  OBJs.append(create_object_2(id=1, name="rack centrifuge", type=1, dimension=struct(length=0, width=0, height=0.106, diameter=0.020), gripper_offset=p[0,0,0.095,0,0,2.356]))
  OBJs.append(create_object_2(id=2, name="sample tube 1", type=2, dimension=struct(length=0, width=0, height=0.106, diameter=0.015), gripper_offset=p[0,0,0,0,0,0]))
  OBJs.append(create_object_2(id=3, name="rack sarstedt", type=3, dimension=struct(length=0, width=0, height=0.100, diameter=0.020), gripper_offset=p[0,0,0,0,0,0]))
  OBJs.append(create_object_2(id=4, name="Lab bottle", type=4, dimension=struct(length=0, width=0, height=0.100, diameter=0.030), gripper_offset=p[0,0,0.2,0,0,0]))
  def create_jig_2(id=0, name="", type=0, capacity=0, jig_offset=p[0,0,0,0,0,0]):
      # iformation about used jigs
      return struct(id=id, name=name, type=type, capacity=capacity, jig_offset=jig_offset)
  end

  JIG2 = create_jig_2()
  JIGs = make_list(0, create_jig_2(), 15)

  JIGs.append(create_jig_2(id=1, name="3FG", type=1, capacity=1, jig_offset=p[0,0,0,0,0,0]))
  JIGs.append(create_jig_2(id=2, name="jig input", type=2, capacity=1, jig_offset=p[0,0,0,0,0,-3.927]))
  JIGs.append(create_jig_2(id=3, name="jig output", type=3, capacity=1, jig_offset=p[0,0,0,0,0,0.78]))
  JIGs.append(create_jig_2(id=6, name="jig bin", type=6, capacity=1, jig_offset=p[0,0,0,0,0,0]))
  JIGs.append(create_jig_2(id=7, name="jig sarstedt racks", type=7, capacity=1, jig_offset=p[0,0,-0.02,0,0,0]))
  JIGs.append(create_jig_2(id=8, name="NoK Bin", type=8, capacity=1, jig_offset=p[0,0,0,0,0,0]))
  JIGs.append(create_jig_2(id=9, name="Pick bott jig", type=9, capacity=1, jig_offset=p[0,0,0,0,0,0]))
  JIGs.append(create_jig_2(id=10, name="Place bott jig", type=10, capacity=1, jig_offset=p[0,0,0,0,0,0]))
  JIGs.append(create_jig_2(id=11, name="bottle shake jig", type=11, capacity=1, jig_offset=p[0,0,0,0,0,0]))
  $ 20 "BeforeStarts"
  $ 21 "uLM"
  $ 22 "CMD_Stop≔ False "
  global CMD_Stop=  False
  $ 23 "CMD_Abort≔ False "
  global CMD_Abort=  False
  $ 24 "CMD_Clear≔ False "
  global CMD_Clear=  False
  $ 25 "STATE≔1"
  global STATE=1
  $ 26 "STATE_Info≔''"
  global STATE_Info=""
  $ 27 "ARM_Referenced≔ False "
  global ARM_Referenced=  False
  $ 28 "zero_ftsensor()"
  zero_ftsensor()
  $ 29 "poses init"
  $ 30 "PSE_A≔p[0,0,0,0,0,0]"
  global PSE_A=p[0,0,0,0,0,0]
  $ 31 "PSE_A_H≔p[0,0,0,0,0,0]"
  global PSE_A_H=p[0,0,0,0,0,0]
  $ 32 "PSE_R≔p[0,0,0,0,0,0]"
  global PSE_R=p[0,0,0,0,0,0]
  $ 33 "PSE_R_H≔p[0,0,0,0,0,0]"
  global PSE_R_H=p[0,0,0,0,0,0]
  $ 34 "PSE_T≔p[0,0,0,0,0,0]"
  global PSE_T=p[0,0,0,0,0,0]
  $ 35 "PSE_T_H≔p[0,0,0,0,0,0]"
  global PSE_T_H=p[0,0,0,0,0,0]
  $ 36 "PSE_C_E≔p[0,0,0,0,0,0]"
  global PSE_C_E=p[0,0,0,0,0,0]
  $ 37 "PSE_C_H≔p[0,0,0,0,0,0]"
  global PSE_C_H=p[0,0,0,0,0,0]
  $ 38 "PSE_C_S≔p[0,0,0,0,0,0]"
  global PSE_C_S=p[0,0,0,0,0,0]
  $ 39 "init_home_by_cartesian_pose(p[0,-0.400,0.300,0,0,0])"
  init_home_by_cartesian_pose(p[0,-0.400,0.300,0,0,0])
  $ 40 "Clearing"
  $ 41 "reset_error()"
  reset_error()
  $ 42 "reset_warning()"
  reset_warning()
  $ 43 "uGo"
  $ 45 "ugo_init( True ,'http://192.168.12.120:10001')"
  ugo_init(  True  ,"http://192.168.12.120:10001")
  $ 46 "ugo_update_outputs()"
  ugo_update_outputs()
  $ 47 "App"
  $ 48 "'ADD APPLICATION SPECIFIC COMMANDS'"
  # 'ADD APPLICATION SPECIFIC COMMANDS'
  $ 49 "Tools"
  $ 50 "OBJ_Picked≔gripper_has_object()"
  global OBJ_Picked=gripper_has_object()
  $ 51 "If OBJ_Picked"
  if (OBJ_Picked):
    # begin: URCap Program Node
    #   Source: Robotiq_Grippers, 1.8.4.4844, Robotiq Inc.
    #   Type: Gripper Activate
    $ 52 "Gripper Activate"

    kill rq_gripper_communication_thread
    rq_gripper_communication_thread_started = False

    rq_init_comm_if_connected(9, "1")
    rq_init_comm_if_connected(2, "2")
    rq_init_comm_if_connected(3, "3")
    rq_init_comm_if_connected(4, "4")
    rq_print_connected_grippers()
    rq_gripper_communication_thread = run rq_gripper_communication()

    while(not rq_gripper_communication_thread_started):
        sync()
    end

    rq_set_max_current_for_all_grippers()

    reset_and_activate = False

    rq_activate_all_grippers(False)
    # end: URCap Program Node
  else:
    $ 53 "Else" "noBreak"
    # begin: URCap Program Node
    #   Source: Robotiq_Grippers, 1.8.4.4844, Robotiq Inc.
    #   Type: Gripper Activate
    $ 54 "Gripper Reset and Activate"

    kill rq_gripper_communication_thread
    rq_gripper_communication_thread_started = False

    rq_init_comm_if_connected(9, "1")
    rq_init_comm_if_connected(2, "2")
    rq_init_comm_if_connected(3, "3")
    rq_init_comm_if_connected(4, "4")
    rq_print_connected_grippers()
    rq_gripper_communication_thread = run rq_gripper_communication()

    while(not rq_gripper_communication_thread_started):
        sync()
    end

    rq_set_max_current_for_all_grippers()

    reset_and_activate = True

    rq_activate_all_grippers(True)
    # end: URCap Program Node
  end
  $ 55 "zero_ftsensor()"
  zero_ftsensor()
  $ 56 "EXTT"
  $ 57 "Set GRP_3F_Enable=Off"
  set_standard_digital_out(4, False)
  $ 58 "Set GRP_3F_Decap=Off"
  set_standard_digital_out(3, False)
  $ 59 "Set GRP_3F_Cap=Off"
  set_standard_digital_out(2, False)
  $ 60 "Set GRP_3F_Open=Off"
  set_standard_digital_out(5, False)
  $ 61 "PSE_T≔get_tool_free_pose(dir=[0,0,0.150], move_in_base_frame=True)"
  global PSE_T=get_tool_free_pose(dir=[0,0,0.150], move_in_base_frame=True)
  $ 62 "If is_reachable(Base_const, [PSE_T])"
  if (is_reachable(p[0.0,0.0,0.0,0.0,0.0,0.0], [PSE_T])):
    $ 63 "MoveL"
    $ 64 "PSE_T" "breakAfter"
    movel(PSE_T, a=1.2, v=0.15)
  end
  while (True):
    $ 65 "Robot Program"
    $ 66 "MAIN"
    $ 67 "command_manager(external_control='uGO', cond_suspend=(ITM_Manipulated and AMR_AtTarget and AMR_Charging and AMR_Battery<40), cond_unsuspend=(AMR_Battery≟60))"
    command_manager(external_control="uGO", cond_suspend=(ITM_Manipulated  and  AMR_AtTarget  and  AMR_Charging  and  AMR_Battery<40), cond_unsuspend=(AMR_Battery == 60))
    $ 68 "log_state(STATE_Info)"
    log_state(STATE_Info)
    $ 69 "Switch STATE"
    switch_1 = STATE
    $ 70 "Case 1"
    if (1 == switch_1):
      $ 71 "Stopping"
      $ 72 "STATE_Info≔'Stopping'"
      global STATE_Info="Stopping"
      $ 73 "end_freedrive_mode()"
      end_freedrive_mode()
      $ 74 "Set"
      set_tcp(p[0.0,0.0,0.161,3.1415,0.0,0.0])
      $ 75 "PSE_T≔get_tool_free_pose(dir=[0,0,0.150], move_in_base_frame=True)"
      global PSE_T=get_tool_free_pose(dir=[0,0,0.150], move_in_base_frame=True)
      $ 76 "If is_reachable(Base_const, [PSE_T])"
      if (is_reachable(p[0.0,0.0,0.0,0.0,0.0,0.0], [PSE_T])):
        $ 77 "MoveL"
        $ 78 "PSE_T" "breakAfter"
        movel(PSE_T, a=1.2, v=0.15)
      end
      $ 79 "do_transition(keep_rxry=OBJ_Picked, r=0)"
      do_transition(keep_rxry=OBJ_Picked, r=0)
      $ 88 "Call Sub_AMR_MiR_V3"
      Sub_AMR_MiR_V3()
      $ 89 "If stopping() and AMR_Done"
      if (stopping()  and  AMR_Done):
        $ 90 "STATE≔2"
        global STATE=2
        $ 91 "ugo_update_outputs()"
        ugo_update_outputs()
      end
    elif (2 == switch_1):
      $ 92 "Case 2"
      $ 93 "Stopped"
      $ 94 "STATE_Info≔'Stopped'"
      global STATE_Info="Stopped"
      $ 95 "Call Sub_AMR_MiR_V3"
      Sub_AMR_MiR_V3()
      $ 96 "If CMD_Reset"
      if (CMD_Reset):
        $ 97 "STATE≔3"
        global STATE=3
        $ 98 "ugo_update_outputs()"
        ugo_update_outputs()
      end
    elif (3 == switch_1):
      $ 99 "Case 3"
      $ 100 " Resetting"
      $ 101 "STATE_Info≔'Resetting'"
      global STATE_Info="Resetting"
      $ 102 "uML"
      $ 103 "reset_error()"
      reset_error()
      $ 104 "reset_warning()"
      reset_warning()
      $ 105 "PROCESS_Step≔0"
      global PROCESS_Step=0
      $ 106 "PROCESS_Info≔''"
      global PROCESS_Info=""
      $ 107 "ARM_Referenced≔ False "
      global ARM_Referenced=  False
      $ 108 "WRK_Done≔ False "
      global WRK_Done=  False
      $ 109 "ITM_Prepared≔ False "
      global ITM_Prepared=  False
      $ 110 "ITM_Manipulated≔ False "
      global ITM_Manipulated=  False
      $ 111 "STP≔0"
      global STP=0
      $ 112 "Action≔0"
      global Action=0
      $ 113 "Action_Info≔''"
      global Action_Info=""
      $ 114 "ITM_ID≔0"
      global ITM_ID=0
      $ 115 "JIG≔0"
      global JIG=0
      $ 116 "JIG_Slot≔0"
      global JIG_Slot=0
      $ 117 "Task_info≔''"
      global Task_info=""
      $ 118 "Set"
      set_tcp(p[0.0,0.0,0.161,3.1415,0.0,0.0])
      $ 119 "App"
      $ 120 "'ADD APPLICATION SPECIFIC COMMANDS'"
      # 'ADD APPLICATION SPECIFIC COMMANDS'
      $ 121 "OBJ_Type≔0"
      global OBJ_Type=0
      $ 122 "OBJ_Nbr≔0"
      global OBJ_Nbr=0
      $ 123 "If CNT_Rack_Output≥50"
      if (CNT_Rack_Output >= 50):
        $ 124 "CNT_Rack_Output≔0"
        global CNT_Rack_Output=0
      end
      $ 125 "TASK≔struct(ID=0, NAVI=struct(target=0, footprint=0, protectiveOff=0, dock=0), WORK=struct(ITM_ID_Src=0, JIG_ID_Src=0, OBJ_Nbr_Src=0, ACT_Src=0, ITM_ID_Tgt=0, JIG_ID_Tgt=0, OBJ_Nbr_Tgt=0, ACT_Tgt=0, OBJ_Type=0))"
      global TASK=struct(ID=0, NAVI=struct(target=0, footprint=0, protectiveOff=0, dock=0), WORK=struct(ITM_ID_Src=0, JIG_ID_Src=0, OBJ_Nbr_Src=0, ACT_Src=0, ITM_ID_Tgt=0, JIG_ID_Tgt=0, OBJ_Nbr_Tgt=0, ACT_Tgt=0, OBJ_Type=0))
      $ 126 "Call Sub_AMR_MiR_V3"
      Sub_AMR_MiR_V3()
      $ 127 "If resetting() and AMR_Done"
      if (resetting()  and  AMR_Done):
        $ 128 "STATE≔4"
        global STATE=4
        $ 129 "ugo_update_outputs()"
        ugo_update_outputs()
      end
    elif (4 == switch_1):
      $ 130 "Case 4"
      $ 131 "Idle"
      $ 132 "STATE_Info≔'Idle'"
      global STATE_Info="Idle"
      $ 133 "If CMD_Start"
      if (CMD_Start):
        $ 134 "STATE≔5"
        global STATE=5
        $ 135 "ugo_update_outputs()"
        ugo_update_outputs()
      end
    elif (5 == switch_1):
      $ 136 "Case 5"
      $ 137 "Starting"
      $ 138 "STATE_Info≔'Starting'"
      global STATE_Info="Starting"
      $ 139 "'ADD COMMANDS WHAT TO START WITH'"
      # 'ADD COMMANDS WHAT TO START WITH'
      $ 140 "Call Sub_AMR_MiR_V3"
      Sub_AMR_MiR_V3()
      $ 141 "get ugo data"
      $ 142 "Assign Tasks"
      $ 143 "TASK.ID = ugo_get_task()"
      TASK.ID = ugo_get_task()
      $ 144 "If TASK.ID≟1"
      if (TASK.ID == 1):
        $ 145 "Task_info≔'Charge'"
        global Task_info="Charge"
        $ 146 "Parameters"
        $ 147 "AMR_PosTarget≔1"
        global AMR_PosTarget=1
      else:
        $ 148 "ElseIf TASK.ID≟9"
        if (TASK.ID == 9):
          $ 149 "'Pick Sarstedt Rack from Variable source'"
          # 'Pick Sarstedt Rack from Variable source'
          $ 150 "Task_info≔'Navigate to Target'"
          global Task_info="Navigate to Target"
          $ 151 "Parameters"
          $ 152 "AMR_PosTarget≔UGO.read_input('00','ITM_ID')"
          global AMR_PosTarget=UGO.read_input("00","ITM_ID")
        else:
          $ 153 "ElseIf TASK.ID≟10"
          if (TASK.ID == 10):
            $ 154 "'Pick Sarstedt Rack from Variable source'"
            # 'Pick Sarstedt Rack from Variable source'
            $ 155 "Task_info≔'Pick Rack'"
            global Task_info="Pick Rack"
            $ 156 "AMR_PosTarget≔2"
            global AMR_PosTarget=2
            $ 157 "Parameters"
            $ 158 "ITM_ID≔UGO.read_input('00','ITM_ID')"
            global ITM_ID=UGO.read_input("00","ITM_ID")
            $ 159 "JIG≔UGO.read_input('00','JIG_ID')"
            global JIG=UGO.read_input("00","JIG_ID")
            $ 160 "OBJ_Type≔3"
            global OBJ_Type=3
          else:
            $ 161 "ElseIf TASK.ID≟11"
            if (TASK.ID == 11):
              $ 162 "'Place Sarstedt Rack on Variable target'"
              # 'Place Sarstedt Rack on Variable target'
              $ 163 "Task_info≔'Place Rack'"
              global Task_info="Place Rack"
              $ 164 "AMR_PosTarget≔2"
              global AMR_PosTarget=2
              $ 165 "Parameters"
              $ 166 "ITM_ID≔UGO.read_input('00','ITM_ID')"
              global ITM_ID=UGO.read_input("00","ITM_ID")
              $ 167 "JIG≔UGO.read_input('00','JIG_ID')"
              global JIG=UGO.read_input("00","JIG_ID")
              $ 168 "OBJ_Type≔3"
              global OBJ_Type=3
            else:
              $ 170 "ElseIf TASK.ID≟12"
              if (TASK.ID == 12):
                $ 171 "Task_info≔'Decapping'"
                global Task_info="Decapping"
                $ 172 "Parameters"
                $ 173 "ITM_ID≔1"
                global ITM_ID=1
                $ 174 "AMR_PosTarget≔AMR_PosActual"
                global AMR_PosTarget=AMR_PosActual
                $ 175 "PRC_TubCounter≔0"
                global PRC_TubCounter=0
              else:
                $ 176 "ElseIf TASK.ID≟13"
                if (TASK.ID == 13):
                  $ 177 "Task_info≔'Empty racks'"
                  global Task_info="Empty racks"
                  $ 178 "Parameters"
                  $ 179 "ITM_ID≔1"
                  global ITM_ID=1
                  $ 180 "AMR_PosTarget≔AMR_PosActual"
                  global AMR_PosTarget=AMR_PosActual
                else:
                  $ 181 "ElseIf TASK.ID≟16"
                  if (TASK.ID == 16):
                    $ 182 "Task_info≔'Decap + Barcode'"
                    global Task_info="Decap + Barcode"
                    $ 183 "Parameters"
                    $ 185 "OBJs_String≔UGO.read_input('00','ObjPos')"
                    global OBJs_String=UGO.read_input("00","ObjPos")
                    $ 186 "OBJs_List≔make_list(length = elements_in_string(OBJs_String), initial_value = -1, capacity = 50)"
                    global OBJs_List=make_list(length = elements_in_string(OBJs_String), initial_value = -1, capacity = 50)
                    $ 187 "OBJs_List≔string_to_list(OBJs_String)"
                    global OBJs_List=string_to_list(OBJs_String)
                    $ 188 "ITM_ID≔1"
                    global ITM_ID=1
                    $ 189 "OBJ_Type≔2"
                    global OBJ_Type=2
                    $ 190 "JIG≔7"
                    global JIG=7
                    $ 191 "AMR_PosTarget≔AMR_PosActual"
                    global AMR_PosTarget=AMR_PosActual
                  else:
                    $ 192 "ElseIf TASK.ID≟99"
                    if (TASK.ID == 99):
                      $ 193 "Task_info≔'Decapping and barcode alignment'"
                      global Task_info="Decapping and barcode alignment"
                      $ 194 "Parameters"
                      $ 195 "PRC_TubNumber≔UGO.read_input('00','TubesNb')"
                      global PRC_TubNumber=UGO.read_input("00","TubesNb")
                      $ 196 "PRC_TubCounter≔0"
                      global PRC_TubCounter=0
                      $ 197 "ITM_ID≔1"
                      global ITM_ID=1
                      $ 198 "AMR_PosTarget≔AMR_PosActual"
                      global AMR_PosTarget=AMR_PosActual
                    else:
                      $ 233 "Else" "noBreak"
                      $ 234 "set_error(ERROR_WRONG_ORDER)"
                      set_error(ERROR_WRONG_ORDER)
                    end
                  end
                end
              end
            end
          end
        end
      end
      $ 235 "test ugo"
      $ 236 "Wait: 0.2"
      sleep(0.2)
      $ 237 "ugo_update_outputs()"
      ugo_update_outputs()
      $ 238 "If starting() and AMR_Done"
      if (starting()  and  AMR_Done):
        $ 239 "log_message(Task_info, 'New Task: ')"
        log_message(Task_info, "New Task: ")
        $ 240 "log_message(to_str(TASK.ID), 'Task_ID: ')"
        log_message(to_str(TASK.ID), "Task_ID: ")
        $ 241 "do_transition(keep_rxry=OBJ_Picked)"
        do_transition(keep_rxry=OBJ_Picked)
        $ 242 "STATE≔6"
        global STATE=6
        $ 243 "ugo_update_outputs()"
        ugo_update_outputs()
      end
    elif (6 == switch_1):
      $ 244 "Case 6"
      $ 245 "Execute"
      $ 246 "STATE_Info≔'Execute'"
      global STATE_Info="Execute"
      $ 247 "If  not CMD_Hold and not CMD_Suspend"
      global thread_flag_247=0
      thread Thread_if_247():
        $ 248 "Switch PROCESS_Step"
        switch_2 = PROCESS_Step
        $ 249 "Case 0"
        if (0 == switch_2):
          $ 250 "PROCESS_Info≔'process control'"
          global PROCESS_Info="process control"
          $ 251 "log_process(PROCESS_Info)"
          log_process(PROCESS_Info)
          $ 252 "process control"
          $ 253 "If  not AMR_AtTarget"
          if (  not  AMR_AtTarget):
            $ 254 "PROCESS_Step≔1"
            global PROCESS_Step=1
          else:
            $ 255 "ElseIf (( not ITM_Prepared and  not WRK_Done) or (ITM_Prepared and WRK_Done))"
            if (((  not  ITM_Prepared  and    not  WRK_Done)  or  (ITM_Prepared  and  WRK_Done))):
              $ 256 "PROCESS_Step≔2"
              global PROCESS_Step=2
            else:
              $ 257 "ElseIf  not WRK_Done"
              if (  not  WRK_Done):
                $ 258 "PROCESS_Step≔3"
                global PROCESS_Step=3
              else:
                $ 259 "Else" "noBreak"
                $ 260 "task finished"
                $ 261 "PROCESS_Info≔''"
                global PROCESS_Info=""
                $ 262 "STATE≔7"
                global STATE=7
                $ 263 "ugo_update_outputs()"
                ugo_update_outputs()
              end
            end
          end
        elif (1 == switch_2):
          $ 264 "Case 1"
          $ 265 "navigate"
          $ 266 "'MOVING THE uML'"
          # 'MOVING THE uML'
          $ 267 "PROCESS_Info≔'move to target'"
          global PROCESS_Info="move to target"
          $ 268 "log_process(PROCESS_Info)"
          log_process(PROCESS_Info)
          $ 269 "If TASK.ID≟1"
          if (TASK.ID == 1):
            $ 270 "Action≔51"
            global Action=51
          else:
            $ 271 "Else" "noBreak"
            $ 272 "Action≔52"
            global Action=52
          end
          $ 273 "Call Sub_AMR_MiR_V3"
          Sub_AMR_MiR_V3()
          $ 274 "If AMR_Done"
          if (AMR_Done):
            $ 275 "PROCESS_Step≔0"
            global PROCESS_Step=0
          end
        elif (2 == switch_2):
          $ 276 "Case 2"
          $ 277 "prepare"
          $ 278 "'THINGS THAT HAVE TO BE DONE ONCE IN A SEQUENCE,WORKFLOW'"
          # 'THINGS THAT HAVE TO BE DONE ONCE IN A SEQUENCE,WORKFLOW'
          $ 279 "PROCESS_Info≔'prepare for work'"
          global PROCESS_Info="prepare for work"
          $ 280 "log_process(PROCESS_Info)"
          log_process(PROCESS_Info)
          $ 281 "If TASK.WORK.ITM_ID_Src>1"
          if (TASK.WORK.ITM_ID_Src>1):
            $ 282 "ITM_ID≔TASK.WORK.ITM_ID_Src"
            global ITM_ID=TASK.WORK.ITM_ID_Src
          else:
            $ 283 "ElseIf TASK.WORK.ITM_ID_Tgt>1"
            if (TASK.WORK.ITM_ID_Tgt>1):
              $ 284 "ITM_ID≔TASK.WORK.ITM_ID_Tgt"
              global ITM_ID=TASK.WORK.ITM_ID_Tgt
            end
          end
          $ 285 "If  not ARM_Referenced and (ITM_ID≠0)"
          if (  not  ARM_Referenced  and  (ITM_ID != 0)):
            $ 286 "STP≔1"
            global STP=1
          else:
            $ 287 "ElseIf ARM_Referenced or (ITM_ID≟0)"
            if (ARM_Referenced  or  (ITM_ID == 0)):
              $ 288 "STP≔2"
              global STP=2
            end
          end
          $ 289 "Switch STP"
          switch_3 = STP
          $ 290 "Case 1"
          if (1 == switch_3):
            $ 291 "reference"
            $ 292 "STP_Info≔'reference at target position'"
            global STP_Info="reference at target position"
            $ 293 "log_step(STP_Info)"
            log_step(STP_Info)
            $ 294 "If ITM_ID≟1"
            if (ITM_ID == 1):
              $ 295 "CAM_Done≔ True "
              global CAM_Done=  True
            else:
              $ 296 "Else" "noBreak"
              $ 297 "Action≔131"
              global Action=131
              $ 298 "Call Sub_Vision_V18"
              Sub_Vision_V18()
            end
            $ 300 "If CAM_Done and  not ERROR.FLAG"
            if (CAM_Done  and    not  ERROR.FLAG):
              $ 301 "log_step('ARM referenced')"
              log_step("ARM referenced")
              $ 302 "ARM_Referenced≔ True "
              global ARM_Referenced=  True
            end
          elif (2 == switch_3):
            $ 303 "Case 2"
            $ 304 "manipulate"
            $ 305 "STP_Info≔'manipulate item'"
            global STP_Info="manipulate item"
            $ 306 "log_step(STP_Info)"
            log_step(STP_Info)
            $ 307 "'In case pressing button is needed'"
            # 'In case pressing button is needed'
            $ 308 "If found_in_list(ITM_ID, ITM_ID_List)"
            if (found_in_list(ITM_ID, ITM_ID_List)):
              $ 309 "Switch ITM_ID"
              switch_4 = ITM_ID
              $ 310 "Case 0"
              if (0 == switch_4):
                $ 311 "ITM_Manipulated≔ not ITM_Manipulated"
                global ITM_Manipulated=  not  ITM_Manipulated
              elif (1 == switch_4):
                $ 312 "Case 1"
                $ 313 "ITM_Manipulated≔ not ITM_Manipulated"
                global ITM_Manipulated=  not  ITM_Manipulated
              elif (2 == switch_4):
                $ 314 "Case 2"
              else:
                $ 324 "Default Case"
                $ 325 "ITM_Manipulated≔ not ITM_Manipulated"
                global ITM_Manipulated=  not  ITM_Manipulated
              end
            end
          end
          $ 326 "ITM_Prepared≔(ITM_Manipulated or  not found_in_list(ITM_ID, ITM_ID_List)) and (ARM_Referenced or ITM_ID≟0) and  not WRK_Done"
          global ITM_Prepared=(ITM_Manipulated  or    not  found_in_list(ITM_ID, ITM_ID_List))  and  (ARM_Referenced  or  ITM_ID == 0)  and    not  WRK_Done
          $ 327 "STP≔0"
          global STP=0
          $ 328 "STP_Info≔''"
          global STP_Info=""
          $ 329 "PROCESS_Step≔0"
          global PROCESS_Step=0
        elif (3 == switch_2):
          $ 330 "Case 3"
          $ 331 "work"
          $ 332 "'ADD EVERY MACHINE, OBJECT, STATION TO WORK ON'"
          # 'ADD EVERY MACHINE, OBJECT, STATION TO WORK ON'
          $ 333 "Switch ITM_ID"
          switch_3 = ITM_ID
          $ 334 "Case 1"
          if (1 == switch_3):
            $ 335 "uLM"
            $ 336 "If TASK.ID≟12"
            if (TASK.ID == 12):
              $ 337 "fill racks"
              $ 338 "Action≔151"
              global Action=151
              $ 339 "Call Sub_Vision_V18"
              Sub_Vision_V18()
              $ 340 "If  not ERROR.FLAG"
              if (  not  ERROR.FLAG):
                $ 341 "Actions for the task"
                $ 342 "Action≔1"
                global Action=1
                $ 343 "JIG≔2"
                global JIG=2
                $ 344 "JIG_Slot≔CAM_Result[0]"
                global JIG_Slot=CAM_Result[0]
                $ 345 "OBJ_Nbr≔CAM_Result[0]"
                global OBJ_Nbr=CAM_Result[0]
                $ 346 "OBJ_Type≔2"
                global OBJ_Type=2
                $ 347 "Call Sub_Action_V4"
                Sub_Action_V4()
                $ 348 "If OBJ_Picked"
                if (OBJ_Picked):
                  $ 349 "CAM_Result.remove(0)"
                  CAM_Result.remove(0)
                  $ 350 "PRC_TubCounter≔PRC_TubCounter+1"
                  global PRC_TubCounter=PRC_TubCounter+1
                  $ 351 "If PRC_TubCounter%4≟0"
                  if (PRC_TubCounter%4 == 0):
                    $ 352 "JIG_Slot≔4"
                    global JIG_Slot=4
                  else:
                    $ 353 "Else" "noBreak"
                    $ 354 "JIG_Slot≔PRC_TubCounter%4"
                    global JIG_Slot=PRC_TubCounter%4
                  end
                  $ 355 "OBJ_Nbr≔ceil(PRC_TubCounter/4)"
                  global OBJ_Nbr=ceil(PRC_TubCounter/4)
                  $ 356 "Action≔2"
                  global Action=2
                  $ 357 "JIG≔4"
                  global JIG=4
                  $ 358 "Call Sub_Action_V4"
                  Sub_Action_V4()
                  $ 359 "Action≔151"
                  global Action=151
                  $ 360 "Call Sub_Vision_V18"
                  Sub_Vision_V18()
                end
              end
              $ 361 "If (CAM_Captures≥CAM_PRM_Retries) or (PRC_TubCounter≥32)"
              if ((CAM_Captures >= CAM_PRM_Retries)  or  (PRC_TubCounter >= 32)):
                $ 362 "PROCESS_Step≔0"
                global PROCESS_Step=0
                $ 363 "WRK_Done≔ True "
                global WRK_Done=  True
              end
            else:
              $ 364 "ElseIf TASK.ID≟10"
              if (TASK.ID == 10):
                $ 365 "Pick Rack"
                $ 366 "Action≔131"
                global Action=131
                $ 367 "Call Sub_Vision_V18"
                Sub_Vision_V18()
                $ 368 "Action≔1"
                global Action=1
                $ 369 "Call Sub_Action_V4"
                Sub_Action_V4()
                $ 370 "PROCESS_Step≔0"
                global PROCESS_Step=0
                $ 371 "WRK_Done≔ True "
                global WRK_Done=  True
              else:
                $ 372 "ElseIf TASK.ID≟11"
                if (TASK.ID == 11):
                  $ 373 "Place Rack"
                  $ 374 "Action≔2"
                  global Action=2
                  $ 375 "Call Sub_Action_V4"
                  Sub_Action_V4()
                  $ 376 "PROCESS_Step≔0"
                  global PROCESS_Step=0
                  $ 377 "WRK_Done≔ True "
                  global WRK_Done=  True
                else:
                  $ 378 "ElseIf TASK.ID≟13"
                  if (TASK.ID == 13):
                    $ 379 "empty racks"
                    $ 380 "pick"
                    $ 381 "Action≔1"
                    global Action=1
                    $ 382 "JIG≔4"
                    global JIG=4
                    $ 383 "If PRC_TubCounter%4≟0"
                    if (PRC_TubCounter%4 == 0):
                      $ 384 "JIG_Slot≔4"
                      global JIG_Slot=4
                    else:
                      $ 385 "Else" "noBreak"
                      $ 386 "JIG_Slot≔PRC_TubCounter%4"
                      global JIG_Slot=PRC_TubCounter%4
                    end
                    $ 387 "OBJ_Nbr≔ceil(PRC_TubCounter/4)"
                    global OBJ_Nbr=ceil(PRC_TubCounter/4)
                    $ 388 "OBJ_Type≔2"
                    global OBJ_Type=2
                    $ 389 "Call Sub_Action_V4"
                    Sub_Action_V4()
                    $ 390 "If OBJ_Picked"
                    if (OBJ_Picked):
                      $ 391 "Action≔2"
                      global Action=2
                      $ 392 "JIG≔3"
                      global JIG=3
                      $ 393 "JIG_Slot≔1"
                      global JIG_Slot=1
                      $ 394 "CNT_Rack_Output≔CNT_Rack_Output + 1"
                      global CNT_Rack_Output=CNT_Rack_Output + 1
                      $ 395 "OBJ_Nbr≔CNT_Rack_Output"
                      global OBJ_Nbr=CNT_Rack_Output
                      $ 396 "Call Sub_Action_V4"
                      Sub_Action_V4()
                      $ 397 "If  not ERROR.FLAG"
                      if (  not  ERROR.FLAG):
                        $ 398 "PRC_TubCounter≔PRC_TubCounter - 1"
                        global PRC_TubCounter=PRC_TubCounter - 1
                      end
                    end
                    $ 399 "If CNT_Rack_Output≥50 or PRC_TubCounter≤0"
                    if (CNT_Rack_Output >= 50  or  PRC_TubCounter <= 0):
                      $ 400 "PROCESS_Step≔0"
                      global PROCESS_Step=0
                      $ 401 "WRK_Done≔ True "
                      global WRK_Done=  True
                    end
                  else:
                    $ 402 "ElseIf TASK.ID≟16"
                    if (TASK.ID == 16):
                      $ 403 "CAM_Result≔OBJs_List"
                      global CAM_Result=OBJs_List
                      $ 404 "PRC_CntDetect≔0"
                      global PRC_CntDetect=0
                      $ 405 "Loop PRC_CntDetect<CAM_Result.length()"
                      while (PRC_CntDetect<CAM_Result.length()):
                        $ 406 "Action≔1"
                        global Action=1
                        $ 407 "ITM_ID≔1"
                        global ITM_ID=1
                        $ 408 "JIG≔2"
                        global JIG=2
                        $ 409 "OBJ_Type≔2"
                        global OBJ_Type=2
                        $ 410 "JIG_Slot≔CAM_Result[PRC_CntDetect]"
                        global JIG_Slot=CAM_Result[PRC_CntDetect]
                        $ 411 "OBJ_Nbr≔CAM_Result[PRC_CntDetect]"
                        global OBJ_Nbr=CAM_Result[PRC_CntDetect]
                        $ 412 "Call Sub_Action_V4"
                        Sub_Action_V4()
                        $ 413 "JIG≔1"
                        global JIG=1
                        $ 414 "Action≔11"
                        global Action=11
                        $ 415 "Call Sub_Action_V4"
                        Sub_Action_V4()
                        $ 416 "Action≔12"
                        global Action=12
                        $ 417 "Call Sub_Action_V4"
                        Sub_Action_V4()
                        $ 418 "Action≔6"
                        global Action=6
                        $ 419 "JIG≔6"
                        global JIG=6
                        $ 420 "Call Sub_Action_V4"
                        Sub_Action_V4()
                        $ 421 "Action≔13"
                        global Action=13
                        $ 422 "Call Sub_Action_V4"
                        Sub_Action_V4()
                        $ 423 "Action≔1"
                        global Action=1
                        $ 424 "JIG≔1"
                        global JIG=1
                        $ 425 "Call Sub_Action_V4"
                        Sub_Action_V4()
                        $ 426 "If OBJ_Brc_OK"
                        if (OBJ_Brc_OK):
                          $ 427 "JIG≔2"
                          global JIG=2
                          $ 428 "Action≔2"
                          global Action=2
                          $ 429 "OBJ_Nbr≔CAM_Result[PRC_CntDetect]"
                          global OBJ_Nbr=CAM_Result[PRC_CntDetect]
                          $ 430 "JIG_Slot≔CAM_Result[PRC_CntDetect]"
                          global JIG_Slot=CAM_Result[PRC_CntDetect]
                          $ 431 "OBJ_Type≔2"
                          global OBJ_Type=2
                          $ 432 "Call Sub_Action_V4"
                          Sub_Action_V4()
                        else:
                          $ 433 "Else" "noBreak"
                          $ 434 "Action≔2"
                          global Action=2
                          $ 435 "JIG≔8"
                          global JIG=8
                          $ 436 "Call Sub_Action_V4"
                          Sub_Action_V4()
                        end
                        $ 437 "PRC_CntDetect≔PRC_CntDetect+1"
                        global PRC_CntDetect=PRC_CntDetect+1
                      end
                      $ 438 "PROCESS_Step≔0"
                      global PROCESS_Step=0
                      $ 439 "WRK_Done≔ True "
                      global WRK_Done=  True
                    end
                  end
                end
              end
            end
          elif (2 == switch_3):
            $ 440 "Case 2"
          elif (5 == switch_3):
            $ 482 "Case 5"
            $ 483 "SarstedtTable"
            $ 484 "Action≔131"
            global Action=131
            $ 485 "Call Sub_Vision_V18"
            Sub_Vision_V18()
            $ 486 "Action≔1"
            global Action=1
            $ 487 "Call Sub_Action_V4"
            Sub_Action_V4()
            $ 488 "PROCESS_Step≔0"
            global PROCESS_Step=0
            $ 489 "WRK_Done≔ True "
            global WRK_Done=  True
          elif (20 == switch_3):
            $ 490 "Case 20"
          else:
            $ 552 "Default Case"
            $ 553 "WRK_Done≔ True "
            global WRK_Done=  True
            $ 554 "PROCESS_Step≔0"
            global PROCESS_Step=0
          end
        end
        thread_flag_247 = 1
      end
      if (  not  CMD_Hold and not CMD_Suspend):
        global thread_handler_247=run Thread_if_247()
        while (thread_flag_247 == 0):
          if not(  not  CMD_Hold and not CMD_Suspend):
            kill thread_handler_247
            thread_flag_247 = 2
          else:
            sync()
          end
        end
      else:
        thread_flag_247 = 2
      end
      $ 555 "If CMD_Hold"
      if (CMD_Hold):
        $ 556 "STATE≔9"
        global STATE=9
        $ 557 "ugo_update_outputs()"
        ugo_update_outputs()
      else:
        $ 558 "ElseIf CMD_Suspend"
        if (CMD_Suspend):
          $ 559 "STATE≔12"
          global STATE=12
          $ 560 "ugo_update_outputs()"
          ugo_update_outputs()
        end
      end
    elif (7 == switch_1):
      $ 561 "Case 7"
      $ 562 "Completing"
      $ 563 "STATE_Info≔'Completing'"
      global STATE_Info="Completing"
      $ 564 "'ADD COMMANDS FOR COMPLETING THE PROCESS'"
      # 'ADD COMMANDS FOR COMPLETING THE PROCESS'
      $ 565 "do_transition(keep_rxry=OBJ_Picked)"
      do_transition(keep_rxry=OBJ_Picked)
      $ 566 "Call Sub_AMR_MiR_V3"
      Sub_AMR_MiR_V3()
      $ 567 "If completing() and AMR_Done"
      if (completing()  and  AMR_Done):
        $ 568 "STATE≔8"
        global STATE=8
        $ 569 "ugo_update_outputs()"
        ugo_update_outputs()
      end
    elif (8 == switch_1):
      $ 570 "Case 8"
      $ 571 "Complete"
      $ 572 "STATE_Info≔'Complete'"
      global STATE_Info="Complete"
      $ 573 "If CMD_Reset"
      if (CMD_Reset):
        $ 574 "STATE≔3"
        global STATE=3
        $ 575 "ugo_update_outputs()"
        ugo_update_outputs()
      end
    elif (9 == switch_1):
      $ 576 "Case 9"
      $ 577 "Holding"
      $ 578 "STATE_Info≔'Holding'"
      global STATE_Info="Holding"
      $ 579 "stopl(0.5)"
      stopl(0.5)
      $ 580 "Call Sub_AMR_MiR_V3"
      Sub_AMR_MiR_V3()
      $ 581 "If holding() and AMR_Done"
      if (holding()  and  AMR_Done):
        $ 582 "STATE≔10"
        global STATE=10
        $ 583 "ugo_update_outputs()"
        ugo_update_outputs()
      end
    elif (10 == switch_1):
      $ 584 "Case 10"
      $ 585 "Held"
      $ 586 "STATE_Info≔'Held'"
      global STATE_Info="Held"
      $ 587 "If CMD_Unhold"
      if (CMD_Unhold):
        $ 588 "end_freedrive_mode()"
        end_freedrive_mode()
        $ 589 "STATE≔11"
        global STATE=11
        $ 590 "ugo_update_outputs()"
        ugo_update_outputs()
      else:
        $ 591 "ElseIf FNC_Freedrive"
        if (FNC_Freedrive):
          $ 592 "freedrive_mode()"
          freedrive_mode()
        else:
          $ 593 "Else" "noBreak"
          $ 594 "end_freedrive_mode()"
          end_freedrive_mode()
        end
      end
    elif (11 == switch_1):
      $ 595 "Case 11"
      $ 596 "Unholding"
      $ 597 "STATE_Info≔'Unholding'"
      global STATE_Info="Unholding"
      $ 598 "Clearing"
      $ 599 "Switch ERROR.ID"
      switch_2 = ERROR.ID
      $ 600 "Case 1002"
      if (1002 == switch_2):
        $ 601 "AMR_AtTarget≔ False "
        global AMR_AtTarget=  False
        $ 602 "ARM_Referenced≔ False "
        global ARM_Referenced=  False
        $ 603 "ITM_Prepared≔ False "
        global ITM_Prepared=  False
        $ 604 "PROCESS_Step≔1"
        global PROCESS_Step=1
      elif (2007 == switch_2):
        $ 605 "Case 2007"
        $ 606 "PROCESS_Step≔1"
        global PROCESS_Step=1
      end
      $ 607 "reset_error()"
      reset_error()
      $ 608 "reset_warning()"
      reset_warning()
      $ 609 "OBJ_Picked≔gripper_has_object()"
      global OBJ_Picked=gripper_has_object()
      $ 610 "Call Sub_AMR_MiR_V3"
      Sub_AMR_MiR_V3()
      $ 611 "If unholding() and AMR_Done"
      if (unholding()  and  AMR_Done):
        $ 612 "STATE≔6"
        global STATE=6
        $ 613 "ugo_update_outputs()"
        ugo_update_outputs()
      end
    elif (12 == switch_1):
      $ 614 "Case 12"
      $ 615 "Suspending"
      $ 616 "STATE_Info≔'Suspending'"
      global STATE_Info="Suspending"
      $ 617 "PROCESS_Info≔str_cat(PROCESS_Info, ' suspended')"
      global PROCESS_Info=str_cat(PROCESS_Info, " suspended")
      $ 618 "If suspending()"
      if (suspending()):
        $ 619 "STATE≔13"
        global STATE=13
        $ 620 "ugo_update_outputs()"
        ugo_update_outputs()
      end
    elif (13 == switch_1):
      $ 621 "Case 13"
      $ 622 "Suspended"
      $ 623 "STATE_Info≔'Suspended'"
      global STATE_Info="Suspended"
      $ 624 "Call Sub_AMR_MiR_V3"
      Sub_AMR_MiR_V3()
      $ 625 "If CMD_Unsuspend"
      if (CMD_Unsuspend):
        $ 626 "STATE≔14"
        global STATE=14
        $ 627 "ugo_update_outputs()"
        ugo_update_outputs()
      end
    elif (14 == switch_1):
      $ 628 "Case 14"
      $ 629 "Unsuspending"
      $ 630 "STATE_Info≔'Unsuspending'"
      global STATE_Info="Unsuspending"
      $ 631 "PROCESS_Step≔0"
      global PROCESS_Step=0
      $ 632 "If unsuspending()"
      if (unsuspending()):
        $ 633 "STATE≔6"
        global STATE=6
        $ 634 "ugo_update_outputs()"
        ugo_update_outputs()
      end
    elif (15 == switch_1):
      $ 635 "Case 15"
      $ 636 "Aborting"
      $ 637 "STATE_Info≔'Aborting'"
      global STATE_Info="Aborting"
      $ 638 "If aborting()"
      if (aborting()):
        $ 639 "STATE≔16"
        global STATE=16
        $ 640 "ugo_update_outputs()"
        ugo_update_outputs()
      end
    elif (16 == switch_1):
      $ 641 "Case 16"
      $ 642 "Aborted"
      $ 643 "STATE_Info≔'Aborted'"
      global STATE_Info="Aborted"
      $ 644 "If CMD_Clear"
      if (CMD_Clear):
        $ 645 "STATE≔17"
        global STATE=17
        $ 646 "ugo_update_outputs()"
        ugo_update_outputs()
      end
    elif (17 == switch_1):
      $ 647 "Case 17"
      $ 648 "Clearing"
      $ 649 "STATE_Info≔'Clearing'"
      global STATE_Info="Clearing"
      $ 650 "Clearing"
      $ 651 "reset_warning()"
      reset_warning()
      $ 652 "reset_error()"
      reset_error()
      $ 653 "If clearing()"
      if (clearing()):
        $ 654 "STATE≔2"
        global STATE=2
        $ 655 "ugo_update_outputs()"
        ugo_update_outputs()
      end
    end
    $ 656 "log_state(STATE_Info)"
    log_state(STATE_Info)
    $ 657 "log_warning(WARNING.MSG)"
    log_warning(WARNING.MSG)
    $ 658 "log_error(ERROR.MSG)"
    log_error(ERROR.MSG)
    $ 659 "Times"
    $ 660 "Switch STATE"
    switch_1 = STATE
    $ 661 "Case 1"
    if (1 == switch_1):
      $ 662 "TM_St_Stopping≔get_time(STATE_Times[STATE-1])"
      global TM_St_Stopping=get_time(STATE_Times[STATE-1])
    elif (2 == switch_1):
      $ 663 "Case 2"
      $ 664 "TM_St_Stopped≔get_time(STATE_Times[STATE-1])"
      global TM_St_Stopped=get_time(STATE_Times[STATE-1])
    elif (3 == switch_1):
      $ 665 "Case 3"
      $ 666 "TM_St_Resetting≔get_time(STATE_Times[STATE-1])"
      global TM_St_Resetting=get_time(STATE_Times[STATE-1])
    elif (4 == switch_1):
      $ 667 "Case 4"
      $ 668 "TM_St_Idle≔get_time(STATE_Times[STATE-1])"
      global TM_St_Idle=get_time(STATE_Times[STATE-1])
    elif (5 == switch_1):
      $ 669 "Case 5"
      $ 670 "TM_St_Starting≔get_time(STATE_Times[STATE-1])"
      global TM_St_Starting=get_time(STATE_Times[STATE-1])
    elif (6 == switch_1):
      $ 671 "Case 6"
      $ 672 "TM_St_Execute≔get_time(STATE_Times[STATE-1])"
      global TM_St_Execute=get_time(STATE_Times[STATE-1])
    elif (7 == switch_1):
      $ 673 "Case 7"
      $ 674 "TM_St_Completin≔get_time(STATE_Times[STATE-1])"
      global TM_St_Completin=get_time(STATE_Times[STATE-1])
    elif (8 == switch_1):
      $ 675 "Case 8"
      $ 676 "TM_St_Complete≔get_time(STATE_Times[STATE-1])"
      global TM_St_Complete=get_time(STATE_Times[STATE-1])
    elif (9 == switch_1):
      $ 677 "Case 9"
      $ 678 "TM_St_Holding≔get_time(STATE_Times[STATE-1])"
      global TM_St_Holding=get_time(STATE_Times[STATE-1])
    elif (10 == switch_1):
      $ 679 "Case 10"
      $ 680 "TM_St_Held≔get_time(STATE_Times[STATE-1])"
      global TM_St_Held=get_time(STATE_Times[STATE-1])
    elif (11 == switch_1):
      $ 681 "Case 11"
      $ 682 "TM_St_Unholding≔get_time(STATE_Times[STATE-1])"
      global TM_St_Unholding=get_time(STATE_Times[STATE-1])
    elif (12 == switch_1):
      $ 683 "Case 12"
      $ 684 "TM_St_Suspendin≔get_time(STATE_Times[STATE-1])"
      global TM_St_Suspendin=get_time(STATE_Times[STATE-1])
    elif (13 == switch_1):
      $ 685 "Case 13"
      $ 686 "TM_St_Suspended≔get_time(STATE_Times[STATE-1])"
      global TM_St_Suspended=get_time(STATE_Times[STATE-1])
    elif (14 == switch_1):
      $ 687 "Case 14"
      $ 688 "TM_St_Unsuspend≔get_time(STATE_Times[STATE-1])"
      global TM_St_Unsuspend=get_time(STATE_Times[STATE-1])
    elif (15 == switch_1):
      $ 689 "Case 15"
      $ 690 "TM_St_Aborting≔get_time(STATE_Times[STATE-1])"
      global TM_St_Aborting=get_time(STATE_Times[STATE-1])
    elif (16 == switch_1):
      $ 691 "Case 16"
      $ 692 "TM_St_Aborted≔get_time(STATE_Times[STATE-1])"
      global TM_St_Aborted=get_time(STATE_Times[STATE-1])
    elif (17 == switch_1):
      $ 693 "Case 17"
      $ 694 "TM_St_Clearing≔get_time(STATE_Times[STATE-1])"
      global TM_St_Clearing=get_time(STATE_Times[STATE-1])
    end
    $ 696 "Wait: 0.1"
    sleep(0.1)
  end
end
